// CONVERTE SECONDI (REAL) IN TIME
FUNCTION F_SecondsToTime : TIME
VAR_INPUT
	rSeconds	:	REAL;
END_VAR
VAR
END_VAR

F_SecondsToTime	:=	REAL_TO_TIME(rSeconds * GVL_Conversions.SECONDS_TO_TIME);

END_FUNCTION

(* stored: Version 1.1.0.1, ProductVersion 3.1.4024.9
   POU F_SecondsToTime: Id {9d168122-d3e8-4d44-b33a-12cef028da27}, SpecialFunc None *)
